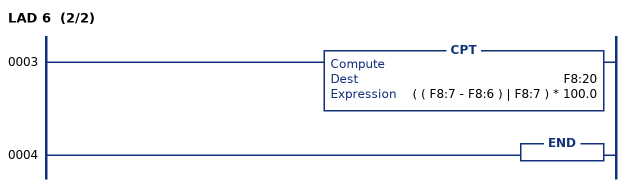
% Rung: 3 %
SOR CPT F8:20 " ( ( F8:7 - F8:6 ) | F8:7 ) * 100.0 " EOR
% Rung: 4 %
SOR END EOR

LADDER 7
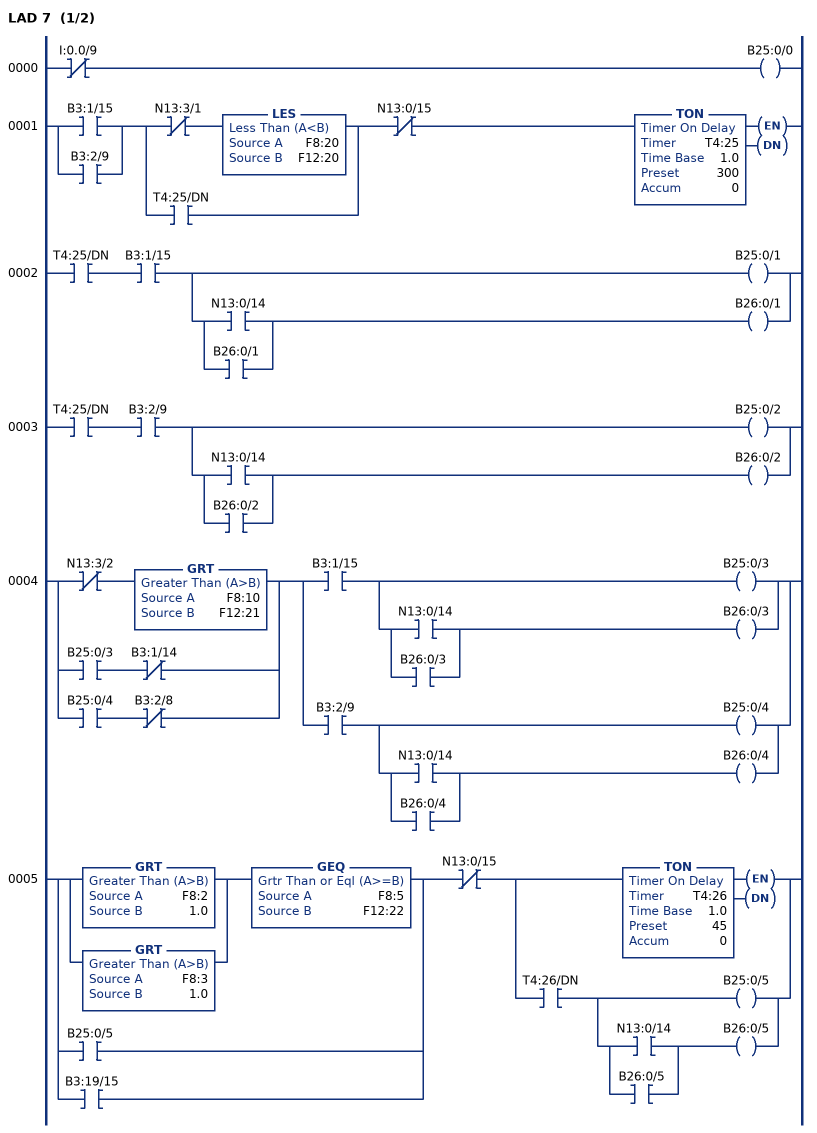
% Rung: 0 %
SOR XIO I:0.0/9 OTE B25:0/0 EOR
% Rung: 1 %
SOR BST XIC B3:1/15 NXB XIC B3:2/9 BND BST XIO N13:3/1 LES F8:20 F12:20 NXB XIC T4:25/DN BND XIO N13:0/15 TON T4:25 1.0 300 0 EOR
% Rung: 2 %
SOR XIC T4:25/DN XIC B3:1/15 BST OTE B25:0/1 NXB BST XIC N13:0/14 NXB XIC B26:0/1 BND OTE B26:0/1 BND EOR
% Rung: 3 %
SOR XIC T4:25/DN XIC B3:2/9 BST OTE B25:0/2 NXB BST XIC N13:0/14 NXB XIC B26:0/2 BND OTE B26:0/2 BND EOR
% Rung: 4 %
SOR BST XIO N13:3/2 GRT F8:10 F12:21 NXB XIC B25:0/3 XIO B3:1/14 NXB XIC B25:0/4 XIO B3:2/8 BND BST XIC B3:1/15 BST OTE B25:0/3 NXB BST XIC N13:0/14 NXB XIC B26:0/3 BND OTE B26:0/3 BND NXB XIC B3:2/9 BST OTE B25:0/4 NXB BST XIC N13:0/14 NXB XIC B26:0/4 BND OTE B26:0/4 BND BND EOR
% Rung: 5 %
SOR BST BST GRT F8:2 1.0 NXB GRT F8:3 1.0 BND GEQ F8:5 F12:22 NXB XIC B25:0/5 NXB XIC B3:19/15 BND XIO N13:0/15 BST TON T4:26 1.0 45 0 NXB XIC T4:26/DN BST OTE B25:0/5 NXB BST XIC N13:0/14 NXB XIC B26:0/5 BND OTE B26:0/5 BND BND EOR

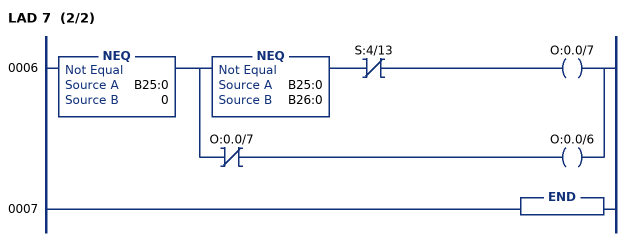
% Rung: 6 %
SOR NEQ B25:0 0 BST NEQ B25:0 B26:0 XIO S:4/13 OTE O:0.0/7 NXB XIO O:0.0/7 OTE O:0.0/6 BND EOR
% Rung: 7 %
SOR END EOR

LADDER 8
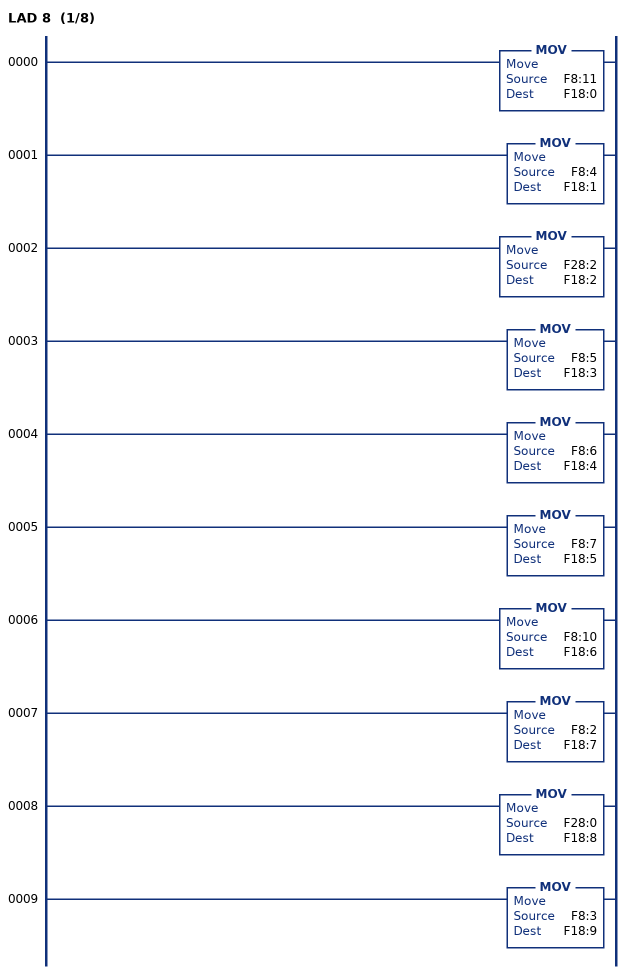
% Rung: 0 %
SOR MOV F8:11 F18:0 EOR
% Rung: 1 %
SOR MOV F8:4 F18:1 EOR
% Rung: 2 %
SOR MOV F28:2 F18:2 EOR
% Rung: 3 %
SOR MOV F8:5 F18:3 EOR
% Rung: 4 %
SOR MOV F8:6 F18:4 EOR
% Rung: 5 %
SOR MOV F8:7 F18:5 EOR
% Rung: 6 %
SOR MOV F8:10 F18:6 EOR
% Rung: 7 %
SOR MOV F8:2 F18:7 EOR
% Rung: 8 %
SOR MOV F28:0 F18:8 EOR
% Rung: 9 %
SOR MOV F8:3 F18:9 EOR

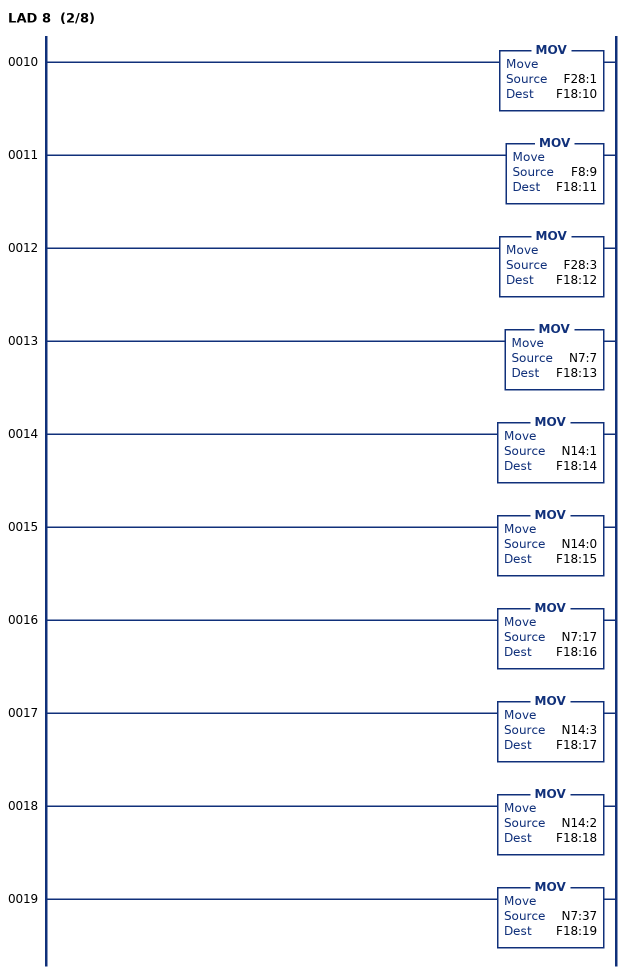
% Rung: 10 %
SOR MOV F28:1 F18:10 EOR
% Rung: 11 %
SOR MOV F8:9 F18:11 EOR
% Rung: 12 %
SOR MOV F28:3 F18:12 EOR
% Rung: 13 %
SOR MOV N7:7 F18:13 EOR
% Rung: 14 %
SOR MOV N14:1 F18:14 EOR
% Rung: 15 %
SOR MOV N14:0 F18:15 EOR
% Rung: 16 %
SOR MOV N7:17 F18:16 EOR
% Rung: 17 %
SOR MOV N14:3 F18:17 EOR
% Rung: 18 %
SOR MOV N14:2 F18:18 EOR
% Rung: 19 %
SOR MOV N7:37 F18:19 EOR

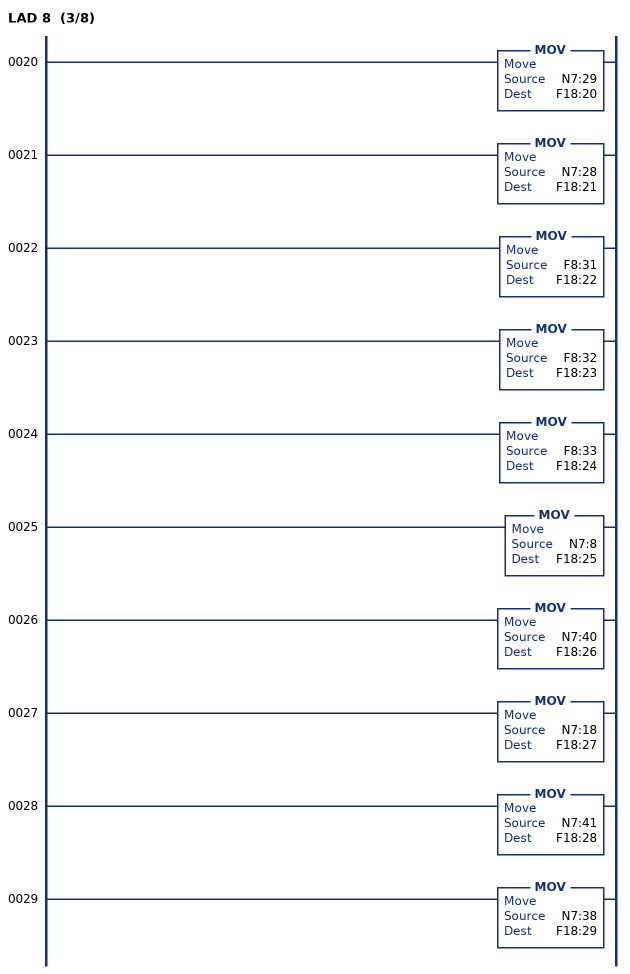
% Rung: 20 %
SOR MOV N7:29 F18:20 EOR
% Rung: 21 %
SOR MOV N7:28 F18:21 EOR
% Rung: 22 %
SOR MOV F8:31 F18:22 EOR
% Rung: 23 %
SOR MOV F8:32 F18:23 EOR
% Rung: 24 %
SOR MOV F8:33 F18:24 EOR
% Rung: 25 %
SOR MOV N7:8 F18:25 EOR
% Rung: 26 %
SOR MOV N7:40 F18:26 EOR
% Rung: 27 %
SOR MOV N7:18 F18:27 EOR
% Rung: 28 %
SOR MOV N7:41 F18:28 EOR
% Rung: 29 %
SOR MOV N7:38 F18:29 EOR

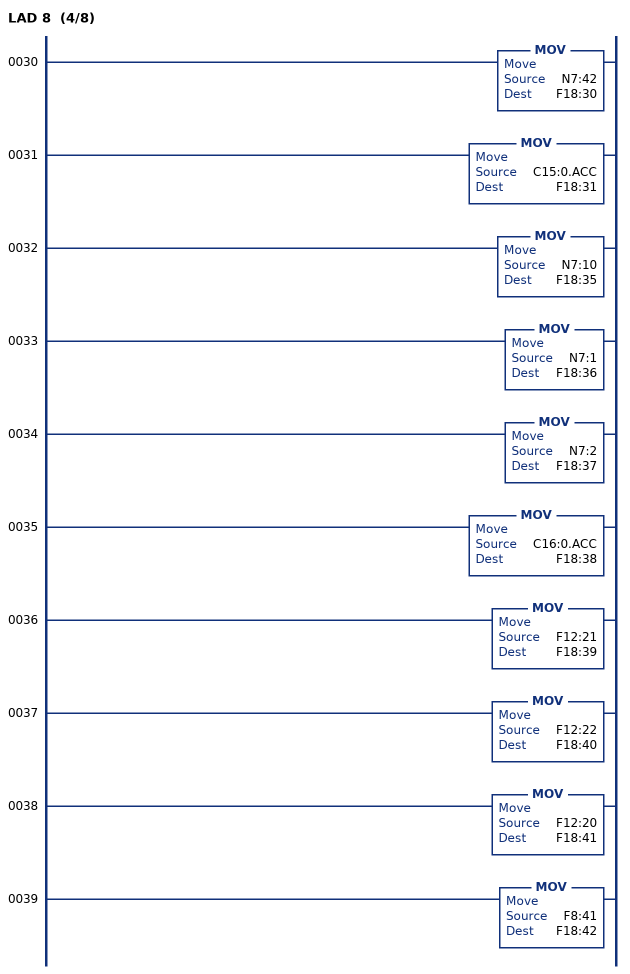
% Rung: 30 %
SOR MOV N7:42 F18:30 EOR
% Rung: 31 %
SOR MOV C15:0.ACC F18:31 EOR
% Rung: 32 %
SOR MOV N7:10 F18:35 EOR
% Rung: 33 %
SOR MOV N7:1 F18:36 EOR
% Rung: 34 %
SOR MOV N7:2 F18:37 EOR
% Rung: 35 %
SOR MOV C16:0.ACC F18:38 EOR
% Rung: 36 %
SOR MOV F12:21 F18:39 EOR
% Rung: 37 %
SOR MOV F12:22 F18:40 EOR
% Rung: 38 %
SOR MOV F12:20 F18:41 EOR
% Rung: 39 %
SOR MOV F8:41 F18:42 EOR

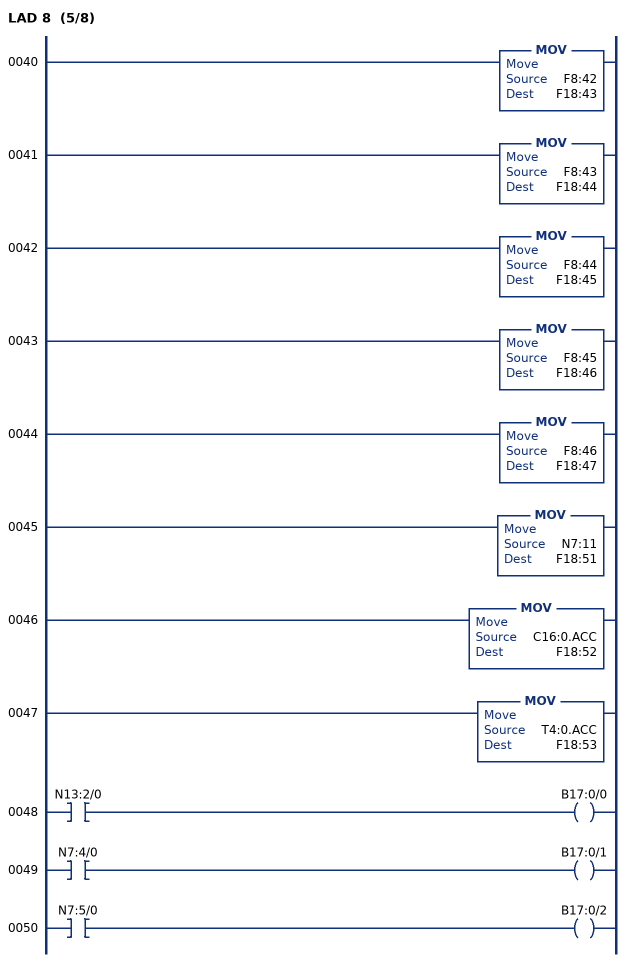
% Rung: 40 %
SOR MOV F8:42 F18:43 EOR
% Rung: 41 %
SOR MOV F8:43 F18:44 EOR
% Rung: 42 %
SOR MOV F8:44 F18:45 EOR
% Rung: 43 %
SOR MOV F8:45 F18:46 EOR
% Rung: 44 %
SOR MOV F8:46 F18:47 EOR
% Rung: 45 %
SOR MOV N7:11 F18:51 EOR
% Rung: 46 %
SOR MOV C16:0.ACC F18:52 EOR
% Rung: 47 %
SOR MOV T4:0.ACC F18:53 EOR
% Rung: 48 %
SOR XIC N13:2/0 OTE B17:0/0 EOR
% Rung: 49 %
SOR XIC N7:4/0 OTE B17:0/1 EOR
% Rung: 50 %
SOR XIC N7:5/0 OTE B17:0/2 EOR

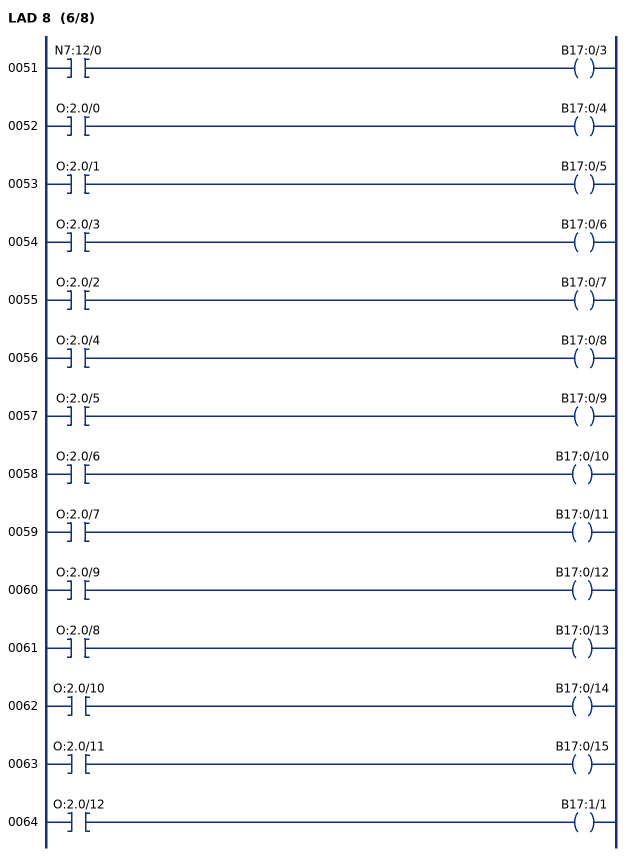
% Rung: 51 %
SOR XIC N7:12/0 OTE B17:0/3 EOR
% Rung: 52 %
SOR XIC O:2.0/0 OTE B17:0/4 EOR
% Rung: 53 %
SOR XIC O:2.0/1 OTE B17:0/5 EOR
% Rung: 54 %
SOR XIC O:2.0/3 OTE B17:0/6 EOR
% Rung: 55 %
SOR XIC O:2.0/2 OTE B17:0/7 EOR
% Rung: 56 %
SOR XIC O:2.0/4 OTE B17:0/8 EOR
% Rung: 57 %
SOR XIC O:2.0/5 OTE B17:0/9 EOR
% Rung: 58 %
SOR XIC O:2.0/6 OTE B17:0/10 EOR
% Rung: 59 %
SOR XIC O:2.0/7 OTE B17:0/11 EOR
% Rung: 60 %
SOR XIC O:2.0/9 OTE B17:0/12 EOR
% Rung: 61 %
SOR XIC O:2.0/8 OTE B17:0/13 EOR
% Rung: 62 %
SOR XIC O:2.0/10 OTE B17:0/14 EOR
% Rung: 63 %
SOR XIC O:2.0/11 OTE B17:0/15 EOR
% Rung: 64 %
SOR XIC O:2.0/12 OTE B17:1/1 EOR

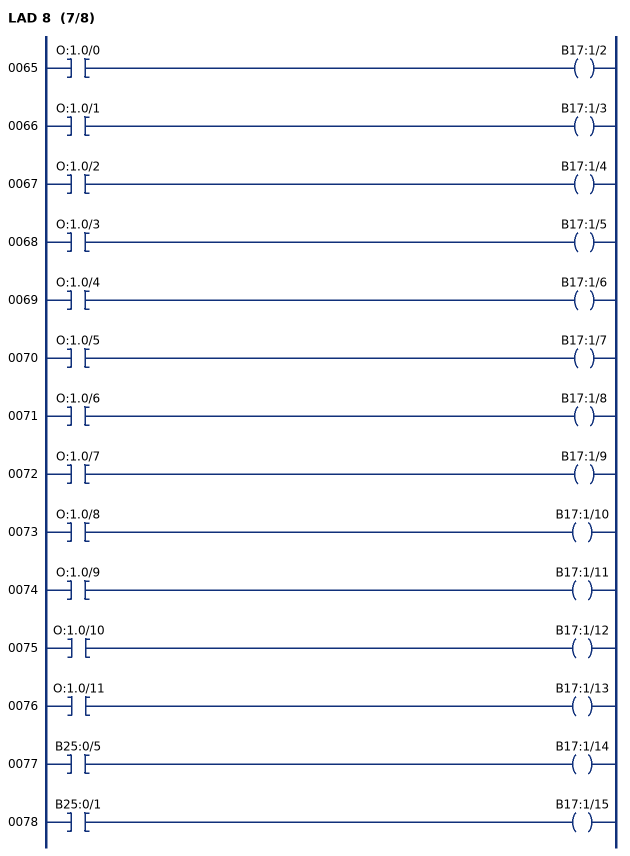
% Rung: 65 %
SOR XIC O:1.0/0 OTE B17:1/2 EOR
% Rung: 66 %
SOR XIC O:1.0/1 OTE B17:1/3 EOR
% Rung: 67 %
SOR XIC O:1.0/2 OTE B17:1/4 EOR
% Rung: 68 %
SOR XIC O:1.0/3 OTE B17:1/5 EOR
% Rung: 69 %
SOR XIC O:1.0/4 OTE B17:1/6 EOR
% Rung: 70 %
SOR XIC O:1.0/5 OTE B17:1/7 EOR
% Rung: 71 %
SOR XIC O:1.0/6 OTE B17:1/8 EOR
% Rung: 72 %
SOR XIC O:1.0/7 OTE B17:1/9 EOR
% Rung: 73 %
SOR XIC O:1.0/8 OTE B17:1/10 EOR
% Rung: 74 %
SOR XIC O:1.0/9 OTE B17:1/11 EOR
% Rung: 75 %
SOR XIC O:1.0/10 OTE B17:1/12 EOR
% Rung: 76 %
SOR XIC O:1.0/11 OTE B17:1/13 EOR
% Rung: 77 %
SOR XIC B25:0/5 OTE B17:1/14 EOR
% Rung: 78 %
SOR XIC B25:0/1 OTE B17:1/15 EOR

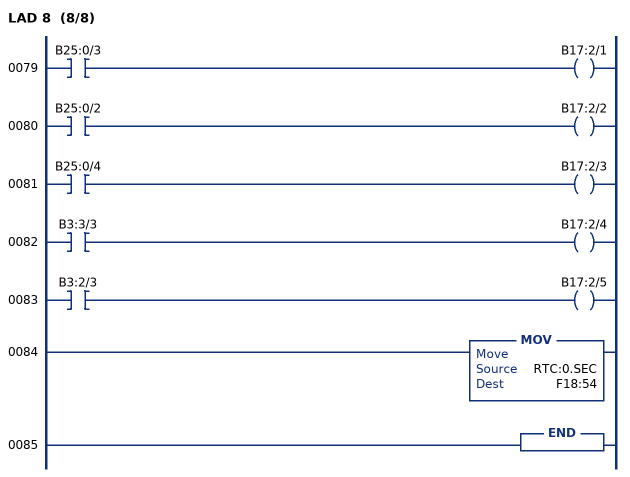
% Rung: 79 %
SOR XIC B25:0/3 OTE B17:2/1 EOR
% Rung: 80 %
SOR XIC B25:0/2 OTE B17:2/2 EOR
% Rung: 81 %
SOR XIC B25:0/4 OTE B17:2/3 EOR
% Rung: 82 %
SOR XIC B3:3/3 OTE B17:2/4 EOR
% Rung: 83 %
SOR XIC B3:2/3 OTE B17:2/5 EOR
% Rung: 84 %
SOR MOV RTC:0.SEC F18:54 EOR
% Rung: 85 %
SOR END EOR

DATA TABLE (non-zero values as saved)
DATA B3
% B3:0 % 0X0000 0X8000 0X0000 0X0400 0X0001 0X0002 0X0000 0X0000 0X0000 0X0000
DATA T4
% .PRE .ACC %
% T4:0 % 15 15
% T4:1 % 1000 160
% T4:2 % 60 0
% T4:3 % 60 0
% T4:9 % 200 0
% T4:10 % 200 0
% T4:11 % 200 0
% T4:12 % 200 0
% T4:13 % 600 0
% T4:15 % 100 37
% T4:20 % 200 0
% T4:21 % 200 0
% T4:22 % 225 0
% T4:23 % 600 0
% T4:25 % 300 0
% T4:26 % 45 0
DATA C5
% .PRE .ACC %
% C5:10 % 2 0
DATA N7
% N7:0 % 0 1 0 1 0 0 1 3 2 9
% N7:10 % 0 0 0 0 0 0 0 3 2 9
% N7:20 % 3 3 3 0 0 150 0 0 5 30
% N7:30 % 0 0 0 0 0 0 0 3 3 3
% N7:40 % 6 6 0 0 0 0 0 0 0 0
DATA F8
% F8:5 % -17.39929 525.3358 550.0611 0 0
% F8:10 % 364.2489 3135.751 0 0 0
% F8:20 % 4.495007 0 0 0 0
% F8:30 % 0 10 5 10 0
% F8:40 % 0 10 35 60 10
% F8:45 % 15 4 0 0 0
DATA N9
% N9:0 % 2025 3 10 1 6 7 14 0 0 1
% N9:10 % 2026 8 24 1 13 4 14
DATA F10
% F10:0 % 1893 2540 2622
DATA F12
% F12:0 % -1000 2000 0 1000 0
% F12:5 % 1000 0 0 0 0
% F12:20 % 0.5 3500 425
DATA N13
% N13:0 % 17 17 1 4 0 4 4 0 0 0
DATA N14
% N14:0 % 5 30 5 30
DATA C15
% .PRE .ACC %
% C15:0 % 4 0
% C15:1 % 100 0
% C15:2 % 50 0
% C15:3 % 100 0
DATA C16
% .PRE .ACC %
% C16:0 % 6 0
% C16:1 % 100 0
% C16:2 % 350 0
% C16:3 % 600 0
% C16:4 % 100 0
% C16:5 % 150 0
% C16:6 % 40 0
DATA B17
% B17:0 % 0X0431 0X00CC 0X0000 0X0000
DATA F18
% F18:0 % 3135.751 0 335.53 -16.48352 525.3358
% F18:5 % 550.3663 364.2489 0 335.53 0
% F18:10 % 335.53 0 335.53 3 30
% F18:15 % 5 3 30 5 3
% F18:20 % 30 5 10 5 10
% F18:25 % 2 6 2 6 3
% F18:35 % 0 1 0 0 3500
% F18:40 % 425 0.5 10 35 60
% F18:45 % 10 15 4 0 0
% F18:50 % 0 0 0 15 14
% F18:55 % 0 58 0 0 0
DATA F19
% F19:0 % 45 0 0 0 0
DATA F28
% F28:0 % 335.53 335.53 335.53 335.53 0
